TYPE T_Percent : LREAL;
END_TYPE

(* stored: Version 1.1.0.1
   DUT T_Percent: Id {4334a5a3-f69e-4772-9496-50776fa5127b} *)
